INTERFACE I_Command

METHOD Start
END_METHOD

METHOD Stop
END_METHOD

METHOD Reset
END_METHOD

METHOD Cycle
VAR_INPUT
    enabled : BOOL;
    sensor : BOOL;
    blocked : BOOL;
END_VAR
END_METHOD

END_INTERFACE

(* stored: Version 1.1.0.1, ProductVersion 3.1 *)
